(* IEC 61131-3 sources: llm-plc-st-eval/data/definitivo/gpt-4o-2024-08-06/B5/zero_shot, 3 files *)

(* ---- ejec_1.st ---- *)
```pascal
FUNCTION_BLOCK FB_Ventilador
VAR
    // Variable de entrada
    quemadorOn : BOOL; // Estado del quemador: TRUE si está encendido, FALSE si está apagado

    // Variable de salida
    ventilador : BOOL; // Estado del ventilador: TRUE si está encendido, FALSE si está apagado

    // Variables internas
    timer : TON; // Temporizador para controlar el tiempo adicional de funcionamiento del ventilador
END_VAR

// Lógica del ventilador
IF quemadorOn THEN
    // Si el quemador está encendido, el ventilador debe estar encendido
    ventilador := TRUE;
    // Reiniciar el temporizador
    timer(IN := FALSE);
ELSE
    // Si el quemador está apagado, iniciar el temporizador
    timer(IN := TRUE, PT := T#30S);
    // El ventilador sigue encendido mientras el temporizador no haya alcanzado el tiempo establecido
    ventilador := timer.Q;
END_IF
END_FUNCTION_BLOCK
```

Este código define un bloque de función `FB_Ventilador` que controla el estado de un ventilador de enfriamiento basado en el estado de un quemador. Utiliza un temporizador `TON` para mantener el ventilador encendido durante 30 segundos adicionales después de que el quemador se apague.

(* ---- ejec_2.st ---- *)
```pascal
FUNCTION_BLOCK FB_Ventilador
VAR
    // Variable de entrada: estado del quemador
    quemadorOn : BOOL;

    // Variable de salida: estado del ventilador
    ventilador : BOOL;

    // Temporizador para controlar el tiempo adicional de funcionamiento del ventilador
    timer : TON;
END_VAR

// Inicialización del temporizador con un tiempo de 30 segundos
timer(IN := NOT quemadorOn, PT := T#30S);

// Lógica para controlar el ventilador
IF quemadorOn THEN
    // Si el quemador está encendido, el ventilador también debe estar encendido
    ventilador := TRUE;
ELSE
    // Si el quemador está apagado, el ventilador sigue encendido hasta que el temporizador expire
    ventilador := NOT timer.Q;
END_IF;

// Actualización del temporizador
timer(IN := NOT quemadorOn);
```

(* ---- ejec_3.st ---- *)
```pascal
FUNCTION_BLOCK FB_Ventilador
VAR
    quemadorOn : BOOL; // Variable de entrada: estado del quemador
    ventilador : BOOL; // Variable de salida: estado del ventilador
    timer : TON; // Temporizador para controlar el tiempo de enfriamiento
END_VAR

// Inicialización del temporizador
timer(IN := FALSE, PT := T#30S);

IF quemadorOn THEN
    // Si el quemador está encendido, el ventilador debe estar encendido
    ventilador := TRUE;
    timer(IN := FALSE); // Asegurarse de que el temporizador esté apagado
ELSE
    // Si el quemador está apagado, iniciar el temporizador
    timer(IN := TRUE);
    IF timer.Q THEN
        // Si el temporizador ha terminado, apagar el ventilador
        ventilador := FALSE;
    ELSE
        // Mientras el temporizador no haya terminado, mantener el ventilador encendido
        ventilador := TRUE;
    END_IF
END_IF
END_FUNCTION_BLOCK
```

Este código define un bloque de función `FB_Ventilador` que controla el estado de un ventilador de enfriamiento basado en el estado de un quemador. Utiliza un temporizador `TON` para mantener el ventilador encendido durante 30 segundos adicionales después de que el quemador se apague.
